(* IEC 61131-3 sources: plc-process-lib/tests/POUs/Suites/FB_Time_Test, 29 files *)

(* ---- BothDelaysOnThenOffTimed.method.decl.st ---- *)
// Обе задержки: включение 1 с, отключение 2 с, шаг 500 мс.
METHOD PRIVATE BothDelaysOnThenOffTimed
VAR
    fbTime  : FB_FakeTime;   // подменное время, старт 1 ч
    fbDelay : FB_Delay;      // ФБ под тестом
END_VAR

(* ---- DelayChangedWhileTimingUsesNewValue.method.decl.st ---- *)
// Изменение задержки во время отсчёта действует сразу: прошедшее время сравнивается с новым
// значением. Уменьшение 10 с → 1 с через 1,5 с — выход в том же вызове; увеличение 2 с → 5 с
// через 1,5 с — выхода нет в 2,0 с и 4,9 с, есть в 5,0 с.
METHOD PRIVATE DelayChangedWhileTimingUsesNewValue
VAR
    fbTime  : FB_FakeTime;   // подменное время, старт 1 ч
    fbShorter : FB_Delay;    // задержку уменьшают
    fbLonger  : FB_Delay;    // задержку увеличивают
    iStep   : INT;           // шаг цикла
END_VAR

(* ---- DelayChangedWhileTimingUsesNewValue.method.impl.st ---- *)
coUnit.TEST('Delay_DelayChangedWhileTiming_UsesNewValue');

fbShorter(xIn := TRUE, tOnDelay := T#10S, itfTime := fbTime);         // t0: фронт
fbLonger(xIn := TRUE, tOnDelay := T#2S, itfTime := fbTime);
FOR iStep := 1 TO 15 DO                                                 // t0 + 1,5 с
    fbTime.Advance(tStep := T#100MS);
    fbShorter(xIn := TRUE, tOnDelay := T#10S, itfTime := fbTime);
    fbLonger(xIn := TRUE, tOnDelay := T#2S, itfTime := fbTime);
END_FOR
fbShorter(xIn := TRUE, tOnDelay := T#1S, itfTime := fbTime);
AssertTrue(Condition := fbShorter.xOut, Message := 'delay reduced below the elapsed time: output at once');
FOR iStep := 1 TO 5 DO                                                  // t0 + 2,0 с
    fbTime.Advance(tStep := T#100MS);
    fbLonger(xIn := TRUE, tOnDelay := T#5S, itfTime := fbTime);
END_FOR
AssertFalse(Condition := fbLonger.xOut, Message := 'delay increased: no output at the old 2 s');
FOR iStep := 1 TO 29 DO                                                 // t0 + 4,9 с
    fbTime.Advance(tStep := T#100MS);
    fbLonger(xIn := TRUE, tOnDelay := T#5S, itfTime := fbTime);
END_FOR
AssertFalse(Condition := fbLonger.xOut, Message := 'no output at t0 + 4.9 s');
fbTime.Advance(tStep := T#100MS);
fbLonger(xIn := TRUE, tOnDelay := T#5S, itfTime := fbTime);             // t0 + 5,0 с
AssertTrue(Condition := fbLonger.xOut, Message := 'output at the new delay 5 s');

coUnit.TEST_FINISHED();

(* ---- FakeTimeAdvanceAddsStep.method.decl.st ---- *)
// Advance прибавляет шаг TIME: два шага по 250 мс, затем длинный шаг 49 сут.
METHOD PRIVATE FakeTimeAdvanceAddsStep
VAR
    fbTime  : FB_FakeTime;   // подменное время, старт 1 ч
    ltMark  : LTIME;         // время перед шагами
END_VAR

(* ---- FakeTimeAdvanceLSubMsAndLongSteps.method.decl.st ---- *)
// AdvanceL: шаги меньше 1 мс (4 по 250 мкс) и больше 49 сут (60 сут).
METHOD PRIVATE FakeTimeAdvanceLSubMsAndLongSteps
VAR
    fbTime  : FB_FakeTime;   // подменное время, старт 1 ч
    ltMark  : LTIME;         // время перед шагами
    iStep   : INT;           // шаг цикла
END_VAR

(* ---- FakeTimeAdvanceLSubMsAndLongSteps.method.impl.st ---- *)
coUnit.TEST('Time_FakeTime_AdvanceL_SubMsAndLongSteps');

ltMark := fbTime.Now();
FOR iStep := 1 TO 4 DO
    fbTime.AdvanceL(ltStep := LTIME#250US);
END_FOR
AssertEquals_LTIME(Expected := LTIME#1MS, Actual := fbTime.Now() - ltMark, Message := 'four steps of 250 us');
ltMark := fbTime.Now();
fbTime.AdvanceL(ltStep := LTIME#60D);
AssertEquals_LTIME(Expected := LTIME#60D, Actual := fbTime.Now() - ltMark, Message := 'LTIME step of 60 days');

coUnit.TEST_FINISHED();

(* ---- FakeTimeSetNowSetsValue.method.decl.st ---- *)
// SetNow ставит время вперёд и назад (назад — допустимо, ФБ библиотеки это переживают).
METHOD PRIVATE FakeTimeSetNowSetsValue
VAR
    fbTime  : FB_FakeTime;   // подменное время, старт 1 ч
END_VAR

(* ---- FakeTimeStartsAtOneHour.method.decl.st ---- *)
// FB_FakeTime стартует с LTIME#1H, а не с 0: ловит код, который считает «0 = не инициализировано».
METHOD PRIVATE FakeTimeStartsAtOneHour
VAR
    fbTime  : FB_FakeTime;   // подменное время, старт 1 ч
END_VAR

(* ---- FakeTimeViaInterfaceReturnsSameTime.method.decl.st ---- *)
// Через I_TimeSource FB_FakeTime отдаёт то же время, что и напрямую (так его получают ФБ библиотеки).
METHOD PRIVATE FakeTimeViaInterfaceReturnsSameTime
VAR
    fbTime  : FB_FakeTime;   // подменное время, старт 1 ч
    itfTime : I_TimeSource;  // источник через интерфейс
END_VAR

(* ---- FirstCallWithInputTrueStartsOnDelay.method.decl.st ---- *)
// Первый вызов сразу с xIn = TRUE ставит отметку и начинает отсчёт. Подменное время стартует с 1 ч:
// без отметки первого вызова разность с нулевой отметкой была бы 1 ч, и выход включился бы сразу.
METHOD PRIVATE FirstCallWithInputTrueStartsOnDelay
VAR
    fbTime  : FB_FakeTime;   // подменное время, старт 1 ч
    fbDelay : FB_Delay;      // ФБ под тестом
END_VAR

(* ---- NoTimeSourceFallsBackToSystemTime.method.decl.st ---- *)
// Без источника (itfTime = 0) FB_Delay берёт встроенный FB_SystemTime: задержка 1 ч идёт и не
// истекает за время теста; нулевая задержка проходит сразу. Реального ожидания нет.
METHOD PRIVATE NoTimeSourceFallsBackToSystemTime
VAR
    fbDelay : FB_Delay;      // задержка 1 ч
    fbZero  : FB_Delay;      // нулевые задержки
END_VAR

(* ---- OffDelayHoldsOutputForDelay.method.decl.st ---- *)
// Задержка отключения 3 с: выход держится до t0 + 2,9 с (идёт отсчёт) и снимается ровно в t0 + 3,0 с.
METHOD PRIVATE OffDelayHoldsOutputForDelay
VAR
    fbTime  : FB_FakeTime;   // подменное время, старт 1 ч
    fbDelay : FB_Delay;      // ФБ под тестом
    iStep   : INT;           // шаг цикла
END_VAR

(* ---- OffDelayHoldsOutputForDelay.method.impl.st ---- *)
coUnit.TEST('Delay_OffDelay_HoldsOutputForDelay');

fbDelay(xIn := TRUE, tOnDelay := T#0S, tOffDelay := T#3S, itfTime := fbTime);
AssertTrue(Condition := fbDelay.xOut, Message := 'zero on-delay: output on at once');
fbDelay(xIn := FALSE, tOnDelay := T#0S, tOffDelay := T#3S, itfTime := fbTime);   // t0: спад
FOR iStep := 1 TO 29 DO
    fbTime.Advance(tStep := T#100MS);
    fbDelay(xIn := FALSE, tOnDelay := T#0S, tOffDelay := T#3S, itfTime := fbTime);
END_FOR
AssertTrue(Condition := fbDelay.xOut, Message := 'output held at t0 + 2.9 s');
AssertTrue(Condition := fbDelay.xTimingOff, Message := 'off-delay timing at t0 + 2.9 s');
fbTime.Advance(tStep := T#100MS);
fbDelay(xIn := FALSE, tOnDelay := T#0S, tOffDelay := T#3S, itfTime := fbTime);   // t0 + 3,0 с
AssertFalse(Condition := fbDelay.xOut, Message := 'output off exactly at t0 + 3.0 s');

coUnit.TEST_FINISHED();

(* ---- OffDelayShortGapIgnored.method.decl.st ---- *)
// Провал входа 1,9 с при задержке отключения 3 с, затем 5 с с TRUE: выход не снимается ни разу.
METHOD PRIVATE OffDelayShortGapIgnored
VAR
    fbTime  : FB_FakeTime;   // подменное время, старт 1 ч
    fbDelay : FB_Delay;      // ФБ под тестом
    iStep   : INT;           // шаг цикла
    xEverOff : BOOL;         // выход снимался хотя бы раз
END_VAR

(* ---- OffDelayShortGapIgnored.method.impl.st ---- *)
coUnit.TEST('Delay_OffDelay_ShortGap_Ignored');

fbDelay(xIn := TRUE, tOffDelay := T#3S, itfTime := fbTime);
fbDelay(xIn := FALSE, tOffDelay := T#3S, itfTime := fbTime);            // t0: спад
xEverOff := NOT fbDelay.xOut;
FOR iStep := 1 TO 19 DO                                                 // вход FALSE до t0 + 1,8 с
    fbTime.Advance(tStep := T#100MS);
    fbDelay(xIn := iStep >= 19, tOffDelay := T#3S, itfTime := fbTime);
    xEverOff := xEverOff OR NOT fbDelay.xOut;
END_FOR
FOR iStep := 1 TO 50 DO
    fbTime.Advance(tStep := T#100MS);
    fbDelay(xIn := TRUE, tOffDelay := T#3S, itfTime := fbTime);
    xEverOff := xEverOff OR NOT fbDelay.xOut;
END_FOR
AssertFalse(Condition := xEverOff, Message := 'gap shorter than the off-delay must be ignored');
AssertFalse(Condition := fbDelay.xTimingOff, Message := 'off-delay timing cancelled');

coUnit.TEST_FINISHED();

(* ---- OnDelayOutputExactlyAtDelay.method.decl.st ---- *)
// Задержка включения 2 с, шаг 100 мс: выход включается ровно на 20-м шаге (t0 + 2,0 с), не на 19-м.
METHOD PRIVATE OnDelayOutputExactlyAtDelay
VAR
    fbTime  : FB_FakeTime;   // подменное время, старт 1 ч
    fbDelay : FB_Delay;      // ФБ под тестом
    iStep   : INT;           // шаг цикла
END_VAR

(* ---- OnDelayOutputExactlyAtDelay.method.impl.st ---- *)
coUnit.TEST('Delay_OnDelay_OutputExactlyAtDelay');

fbDelay(xIn := TRUE, tOnDelay := T#2S, itfTime := fbTime);              // t0: фронт
FOR iStep := 1 TO 19 DO
    fbTime.Advance(tStep := T#100MS);
    fbDelay(xIn := TRUE, tOnDelay := T#2S, itfTime := fbTime);
END_FOR
AssertFalse(Condition := fbDelay.xOut, Message := 'no output at t0 + 1.9 s');
fbTime.Advance(tStep := T#100MS);
fbDelay(xIn := TRUE, tOnDelay := T#2S, itfTime := fbTime);              // t0 + 2,0 с
AssertTrue(Condition := fbDelay.xOut, Message := 'output exactly at t0 + 2.0 s');

coUnit.TEST_FINISHED();

(* ---- OnDelayShortPulseIgnored.method.decl.st ---- *)
// Импульс 1,5 с при задержке включения 2 с, затем 5 с покоя: выход не включается ни разу,
// ожидание отменяется.
METHOD PRIVATE OnDelayShortPulseIgnored
VAR
    fbTime  : FB_FakeTime;   // подменное время, старт 1 ч
    fbDelay : FB_Delay;      // ФБ под тестом
    iStep   : INT;           // шаг цикла
    xEverOn : BOOL;          // выход включался хотя бы раз
END_VAR

(* ---- OnDelayShortPulseIgnored.method.impl.st ---- *)
coUnit.TEST('Delay_OnDelay_ShortPulse_Ignored');

fbDelay(xIn := TRUE, tOnDelay := T#2S, itfTime := fbTime);              // t0: фронт
FOR iStep := 1 TO 15 DO                                                 // вход TRUE до t0 + 1,4 с
    fbTime.Advance(tStep := T#100MS);
    fbDelay(xIn := iStep < 15, tOnDelay := T#2S, itfTime := fbTime);
    xEverOn := xEverOn OR fbDelay.xOut;
END_FOR
FOR iStep := 1 TO 50 DO
    fbTime.Advance(tStep := T#100MS);
    fbDelay(xIn := FALSE, tOnDelay := T#2S, itfTime := fbTime);
    xEverOn := xEverOn OR fbDelay.xOut;
END_FOR
AssertFalse(Condition := xEverOn, Message := 'pulse shorter than the on-delay must be ignored');
AssertFalse(Condition := fbDelay.xTimingOn, Message := 'timing must be cancelled when the input returns');

coUnit.TEST_FINISHED();

(* ---- PresetForcesOutputWithoutDelay.method.decl.st ---- *)
// Preset ставит выход сразу, без задержек включения и отключения (5 с каждая).
METHOD PRIVATE PresetForcesOutputWithoutDelay
VAR
    fbTime  : FB_FakeTime;   // подменное время, старт 1 ч
    fbDelay : FB_Delay;      // ФБ под тестом
END_VAR

(* ---- PresetRestartsTimingOnNextCall.method.decl.st ---- *)
// После Preset отсчёт начинается заново с ближайшего вызова тела: задержка 2 с, через 1,5 с
// Preset(FALSE), следующий вызов в t0 + 1,6 с — выход только в t0 + 3,6 с, а не в t0 + 2,0 с.
METHOD PRIVATE PresetRestartsTimingOnNextCall
VAR
    fbTime  : FB_FakeTime;   // подменное время, старт 1 ч
    fbDelay : FB_Delay;      // ФБ под тестом
    iStep   : INT;           // шаг цикла
END_VAR

(* ---- PresetRestartsTimingOnNextCall.method.impl.st ---- *)
coUnit.TEST('Delay_Preset_RestartsTimingOnNextCall');

fbDelay(xIn := TRUE, tOnDelay := T#2S, itfTime := fbTime);              // t0: фронт
FOR iStep := 1 TO 15 DO                                                 // t0 + 1,5 с
    fbTime.Advance(tStep := T#100MS);
    fbDelay(xIn := TRUE, tOnDelay := T#2S, itfTime := fbTime);
END_FOR
fbDelay.Preset(xValue := FALSE);
FOR iStep := 1 TO 5 DO                                                  // t0 + 1,6 с — новая отметка
    fbTime.Advance(tStep := T#100MS);                                   // ... t0 + 2,0 с
    fbDelay(xIn := TRUE, tOnDelay := T#2S, itfTime := fbTime);
END_FOR
AssertFalse(Condition := fbDelay.xOut, Message := 'old timing must not complete after Preset');
FOR iStep := 1 TO 15 DO                                                 // t0 + 3,5 с
    fbTime.Advance(tStep := T#100MS);
    fbDelay(xIn := TRUE, tOnDelay := T#2S, itfTime := fbTime);
END_FOR
AssertFalse(Condition := fbDelay.xOut, Message := 'no output 1.9 s after the restart');
fbTime.Advance(tStep := T#100MS);
fbDelay(xIn := TRUE, tOnDelay := T#2S, itfTime := fbTime);              // t0 + 3,6 с
AssertTrue(Condition := fbDelay.xOut, Message := 'output 2.0 s after the restart');

coUnit.TEST_FINISHED();

(* ---- RemainingReportsTimeLeft.method.decl.st ---- *)
// tRemaining: полная задержка сразу после фронта, остаток по ходу отсчёта, T#0S без отсчёта;
// то же для задержки отключения.
METHOD PRIVATE RemainingReportsTimeLeft
VAR
    fbTime  : FB_FakeTime;   // подменное время, старт 1 ч
    fbDelay : FB_Delay;      // ФБ под тестом
END_VAR

(* ---- SystemTimeIsMonotonic.method.decl.st ---- *)
// Дымовая проверка FB_SystemTime (оператор LTIME()): 20 000 вызовов подряд — время не убывает,
// растёт (значит, берётся заново в каждом вызове) и больше нуля. Реального ожидания нет.
// Проверка R1 контракта; ручная проверка со сменой времени ОС — docs/MANUAL_STEPS.md.
METHOD PRIVATE SystemTimeIsMonotonic
VAR
    fbSys      : FB_SystemTime;   // ФБ под тестом
    itfTime    : I_TimeSource;    // через интерфейс, как в ФБ библиотеки
    ltFirst    : LTIME;           // время первого вызова
    ltPrev     : LTIME;           // время предыдущего вызова
    ltNow      : LTIME;           // время этого вызова
    xMonotonic : BOOL := TRUE;    // ни разу не убывало
    iStep      : INT;             // шаг цикла
END_VAR

(* ---- SystemTimeIsMonotonic.method.impl.st ---- *)
coUnit.TEST('Time_SystemTime_IsMonotonic');

itfTime := fbSys;
ltFirst := itfTime.Now();
ltPrev := ltFirst;
FOR iStep := 1 TO 20000 DO
    ltNow := itfTime.Now();
    xMonotonic := xMonotonic AND (ltNow >= ltPrev);
    ltPrev := ltNow;
END_FOR
AssertTrue(Condition := xMonotonic, Message := 'LTIME() must not decrease over 20000 calls');
AssertTrue(Condition := ltPrev > ltFirst, Message := 'system time must advance from call to call');
AssertTrue(Condition := ltFirst > LTIME#0S, Message := 'system time must be above zero');

coUnit.TEST_FINISHED();

(* ---- TimeGoesBackwardsRestartsTiming.method.decl.st ---- *)
// «Время назад» (SetNow на 11,5 с раньше) во время отсчёта: выход не меняется, остаток — полная
// задержка (разность LTIME без переполнения), выход ровно через 2 с от нового времени.
METHOD PRIVATE TimeGoesBackwardsRestartsTiming
VAR
    fbTime  : FB_FakeTime;   // подменное время, старт 1 ч
    fbDelay : FB_Delay;      // ФБ под тестом
    iStep   : INT;           // шаг цикла
END_VAR

(* ---- TimeGoesBackwardsRestartsTiming.method.impl.st ---- *)
coUnit.TEST('Delay_TimeGoesBackwards_RestartsTiming');

fbDelay(xIn := TRUE, tOnDelay := T#2S, itfTime := fbTime);              // t0 = 1 ч
FOR iStep := 1 TO 15 DO                                                 // t0 + 1,5 с
    fbTime.Advance(tStep := T#100MS);
    fbDelay(xIn := TRUE, tOnDelay := T#2S, itfTime := fbTime);
END_FOR
fbTime.SetNow(ltValue := LTIME#59M50S);                                 // назад на 11,5 с
fbDelay(xIn := TRUE, tOnDelay := T#2S, itfTime := fbTime);
AssertFalse(Condition := fbDelay.xOut, Message := 'time going backwards must not switch the output');
AssertEquals_TIME(Expected := T#2S, Actual := fbDelay.tRemaining,
                  Message := 'timing restarts with the full delay, no unsigned overflow');
FOR iStep := 1 TO 19 DO
    fbTime.Advance(tStep := T#100MS);
    fbDelay(xIn := TRUE, tOnDelay := T#2S, itfTime := fbTime);
END_FOR
AssertFalse(Condition := fbDelay.xOut, Message := 'no output 1.9 s after the restart');
fbTime.Advance(tStep := T#100MS);
fbDelay(xIn := TRUE, tOnDelay := T#2S, itfTime := fbTime);
AssertTrue(Condition := fbDelay.xOut, Message := 'output 2.0 s after the restart');

coUnit.TEST_FINISHED();

(* ---- TimingFlagsReflectCountdown.method.decl.st ---- *)
// xTimingOn и xTimingOff взведены только во время своих отсчётов (задержки по 1 с).
METHOD PRIVATE TimingFlagsReflectCountdown
VAR
    fbTime  : FB_FakeTime;   // подменное время, старт 1 ч
    fbDelay : FB_Delay;      // ФБ под тестом
END_VAR

(* ---- ZeroDelaysPassThroughSameCall.method.decl.st ---- *)
// Задержки T#0S: фронт и спад проходят в том же вызове, отсчёта нет. Время не продвигается.
METHOD PRIVATE ZeroDelaysPassThroughSameCall
VAR
    fbTime  : FB_FakeTime;   // подменное время, старт 1 ч
    fbDelay : FB_Delay;      // ФБ под тестом
END_VAR
